// Mitsubishi GX Works2 project: FX2N   PLC: FX2N/FX2NC

PROGRAM MAIN
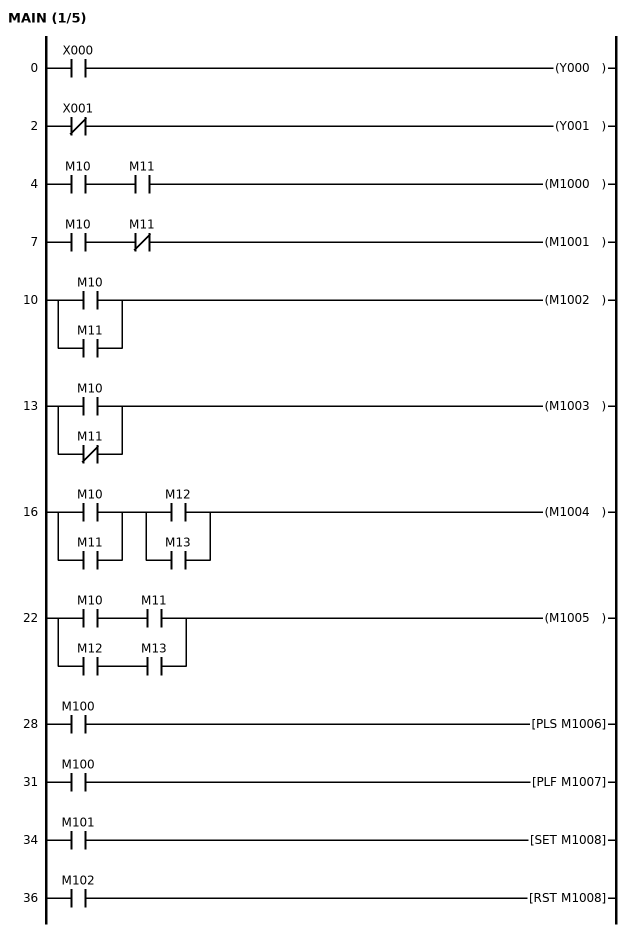
0     LD      X000
      OUT     Y000
2     LDI     X001
      OUT     Y001
4     LD      M10
      AND     M11
      OUT     M1000
7     LD      M10
      ANI     M11
      OUT     M1001
10    LD      M10
      OR      M11
      OUT     M1002
13    LD      M10
      ORI     M11
      OUT     M1003
16    LD      M10
      OR      M11
      LD      M12
      OR      M13
      ANB
      OUT     M1004
22    LD      M10
      AND     M11
      LD      M12
      AND     M13
      ORB
      OUT     M1005
28    LD      M100
      PLS     M1006
31    LD      M100
      PLF     M1007
34    LD      M101
      SET     M1008
36    LD      M102
      RST     M1008
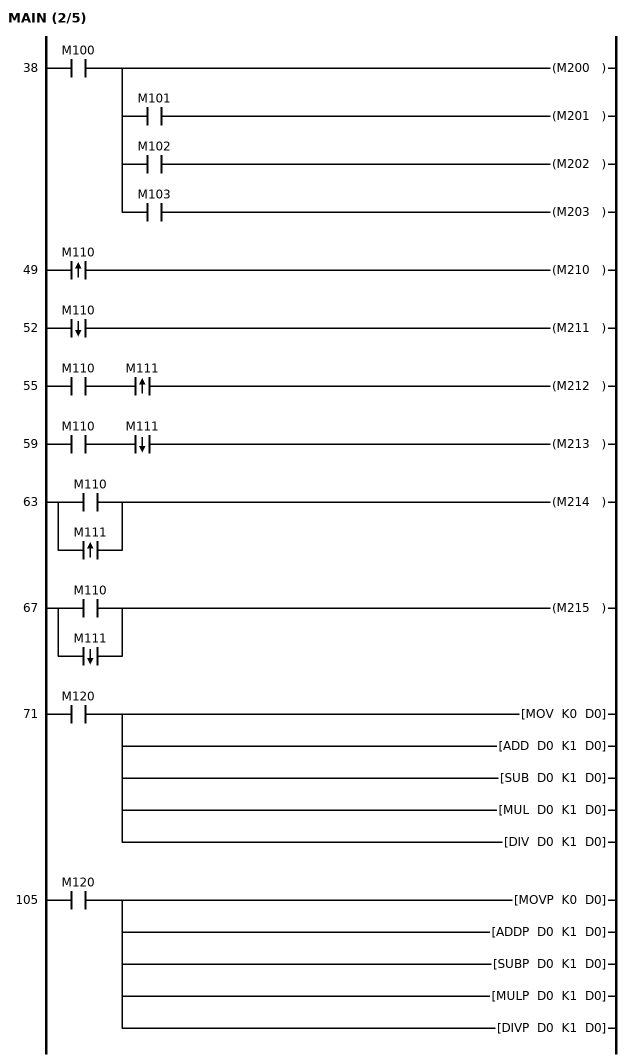
38    LD      M100
      OUT     M200
      MPS
      AND     M101
      OUT     M201
      MRD
      AND     M102
      OUT     M202
      MPP
      AND     M103
      OUT     M203
49    LDP     M110
      OUT     M210
52    LDF     M110
      OUT     M211
55    LD      M110
      ANDP    M111
      OUT     M212
59    LD      M110
      ANDF    M111
      OUT     M213
63    LD      M110
      ORP     M111
      OUT     M214
67    LD      M110
      ORF     M111
      OUT     M215
71    LD      M120
      MOV     K0 D0
      ADD     D0 K1 D0
      SUB     D0 K1 D0
      MUL     D0 K1 D0
      DIV     D0 K1 D0
105   LD      M120
      MOVP    K0 D0
      ADDP    D0 K1 D0
      SUBP    D0 K1 D0
      MULP    D0 K1 D0
      DIVP    D0 K1 D0
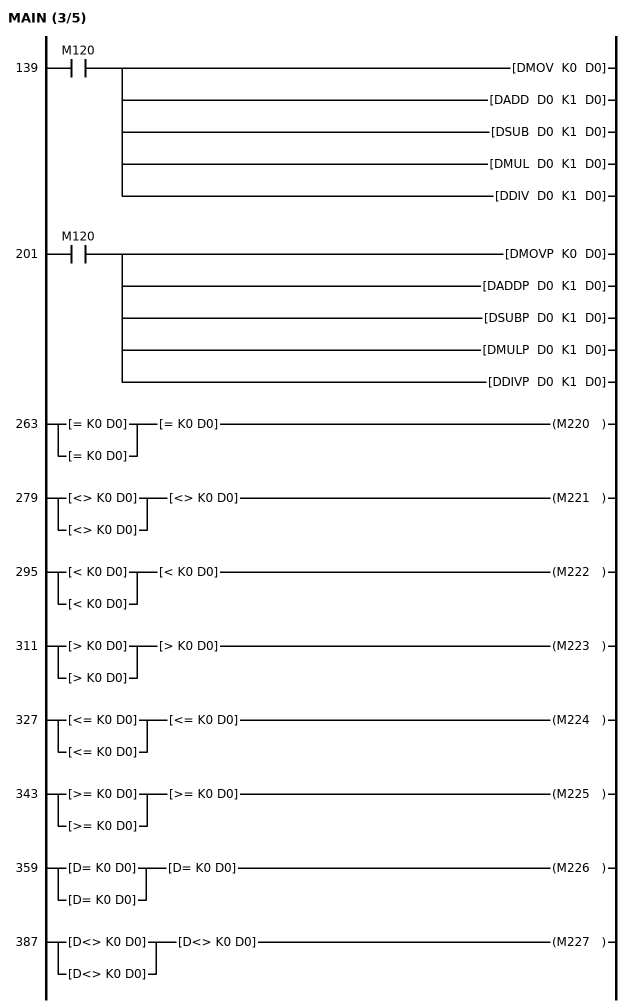
139   LD      M120
      DMOV    K0 D0
      DADD    D0 K1 D0
      DSUB    D0 K1 D0
      DMUL    D0 K1 D0
      DDIV    D0 K1 D0
201   LD      M120
      DMOVP   K0 D0
      DADDP   D0 K1 D0
      DSUBP   D0 K1 D0
      DMULP   D0 K1 D0
      DDIVP   D0 K1 D0
263   LD=     K0 D0
      OR=     K0 D0
      AND=    K0 D0
      OUT     M220
279   LD<>    K0 D0
      OR<>    K0 D0
      AND<>   K0 D0
      OUT     M221
295   LD<     K0 D0
      OR<     K0 D0
      AND<    K0 D0
      OUT     M222
311   LD>     K0 D0
      OR>     K0 D0
      AND>    K0 D0
      OUT     M223
327   LD<=    K0 D0
      OR<=    K0 D0
      AND<=   K0 D0
      OUT     M224
343   LD>=    K0 D0
      OR>=    K0 D0
      AND>=   K0 D0
      OUT     M225
359   LDD=    K0 D0
      ORD=    K0 D0
      ANDD=   K0 D0
      OUT     M226
387   LDD<>   K0 D0
      ORD<>   K0 D0
      ANDD<>  K0 D0
      OUT     M227
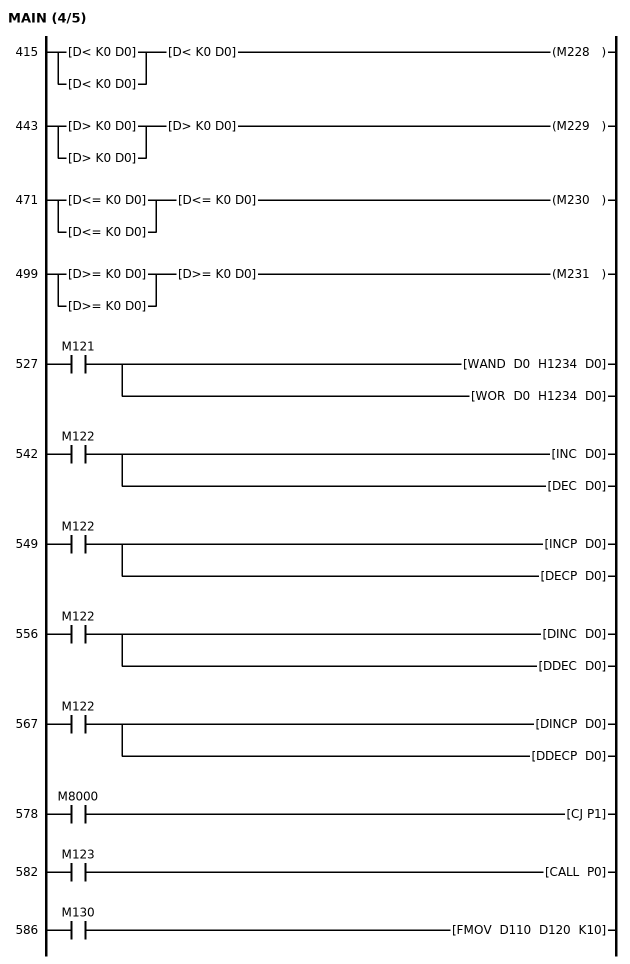
415   LDD<    K0 D0
      ORD<    K0 D0
      ANDD<   K0 D0
      OUT     M228
443   LDD>    K0 D0
      ORD>    K0 D0
      ANDD>   K0 D0
      OUT     M229
471   LDD<=   K0 D0
      ORD<=   K0 D0
      ANDD<=  K0 D0
      OUT     M230
499   LDD>=   K0 D0
      ORD>=   K0 D0
      ANDD>=  K0 D0
      OUT     M231
527   LD      M121
      WAND    D0 H1234 D0
      WOR     D0 H1234 D0
542   LD      M122
      INC     D0
      DEC     D0
549   LD      M122
      INCP    D0
      DECP    D0
556   LD      M122
      DINC    D0
      DDEC    D0
567   LD      M122
      DINCP   D0
      DDECP   D0
578   LD      M8000
      CJ      P1
582   LD      M123
      CALL    P0
586   LD      M130
      FMOV    D110 D120 K10
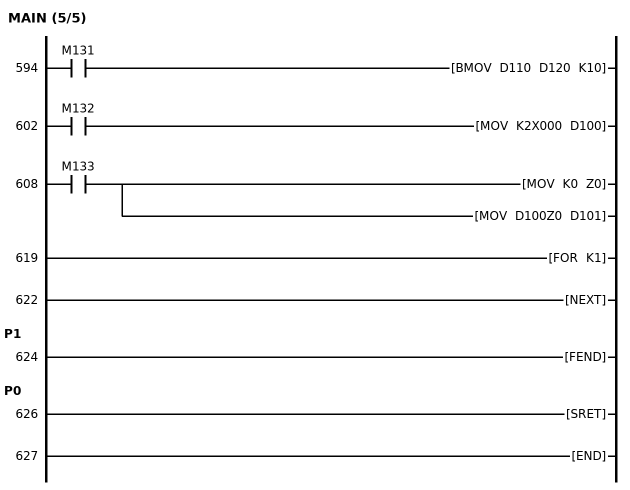
594   LD      M131
      BMOV    D110 D120 K10
602   LD      M132
      MOV     K2X000 D100
608   LD      M133
      MOV     K0 Z0
      MOV     D100Z0 D101
619   FOR     K1
622   NEXT
      P1
624   FEND
      P0
626   SRET
627   END
END_PROGRAM
